(* Schneider Machine Expert - Basic project Projeto Sharpy 2 - Encoder e botão, file version 3.0.0.0 *)
(* ProjectInformations: Name=Novo projeto *)

HARDWARE
  Cpu 0: TM221CE40R
  EthernetConfiguration: NetworkName=M221, IpAllocationMode=FixedAddress, IpAddress=10.0.0.20, SubnetMask=255.0.0.0
  SerialLineConfiguration: Baud=Baud19200, Parity=ParityEven, DataBits=DataBits8, StopBits=StopBits1, PhysicalMedium=PhysicalMediumRs485, TransmissionMode=TransmissionModeModbusRtu, SlaveId=1, Addressing=SlaveAddressing
  MastTask: UsePeriodScanMode=false, PeriodScan=100
  FastTask: Period=255
  CpuBehavior: StartingMode=StartAsPreviousState, AutoSaveRamOnEeprom=true, WatchdogPeriod=250

SYMBOLS  (address, symbol, comment, settings)
  %HSC0.V   VALOR_ENCODER  "Entrada de alta velocidade"
  %S6       SB_TB1S  "Base de tempo de 1 s gerada por um relógio interno"
  %MW0      PULSOS_ENCODER  "Pulsos brutos do encoder"
  %MF2      ANGULO_ATUAL  "Ângulo instantâneo em Graus"
  %MF4      ANGULO_PICO  "Maior ângulo atingido no impacto"
  %MF6      ENERGIA_NOMINAL  "Capacidade da ponta do martelo"
  %MF8      ENERGIA_ABSORVIDA  "Resultado final do ensaio em Joules"
  %MF10     MF_10
  %MF12     MF_12
  %TM0        [Type=TP, Preset=7, Base=OneSecond]
  %TM1        [Type=TP, Preset=7, Base=OneSecond]
  %TM2        [Type=TP, Preset=7, Base=OneSecond]
  %I0.2     BOT_RESET  "Botão físico de zerar encoder e pico"
  %I0.17    SENSOR_PORTA  "Sensor se a porta está fechada"
  %I0.18    SENSOR_BAIXO  "Sensor se o braço está em cima"
  %I0.19    SENSOR_CIMA  "Sensor se o braço está em cima"
  %I0.20    BOTÃO_ZERAR
  %I0.21    BOTÃO_IMPACTO  "Botão que libera para o impacto"
  %I0.22    BOTÃO_DESCER  "Botão que aciona por 7s"
  %I0.23    BOTÃO_SUBIR  "Botão que aciona por 7s"
  %Q0.0       "Motor Descer"
  %Q0.1       "Motor Subir"
  %Q0.2       "Disparo impacto"
  %Q0.3     Q_0_3
  %Q0.4     Q_0_4
  %Q0.5     Q_0_5
  %Q0.14    Q_0_14
  %Q0.15    Q_0_15  "Led porta"
  %IW0.0    IN_ANALOG  "Valor do Potenciômetro"  [Type=Type_0_10V, Scope=Scope_Normal, Minimum=0, Maximum=1000]
  %HSC0       [Type=CounterOrDownCounterBiPhasesX4, Preset=0, DedicatedInputs(DedicatedInput(Activated=true), DedicatedInput(Activated=true)), ReflexOutputs(ReflexOutput(Activated=false, LessThanS0=false, GreaterOrEqualThanS0=false, GreaterOrEqualThanS1=false), ReflexOutput(Activated=false, LessThanS0=false, GreaterOrEqualThanS0=false, GreaterOrEqualThanS1=false)), Thresholds(Threshold(ThresholdType=NotUsed, Pri]

POU Novo POU
  (* SectionNumber=1 *)

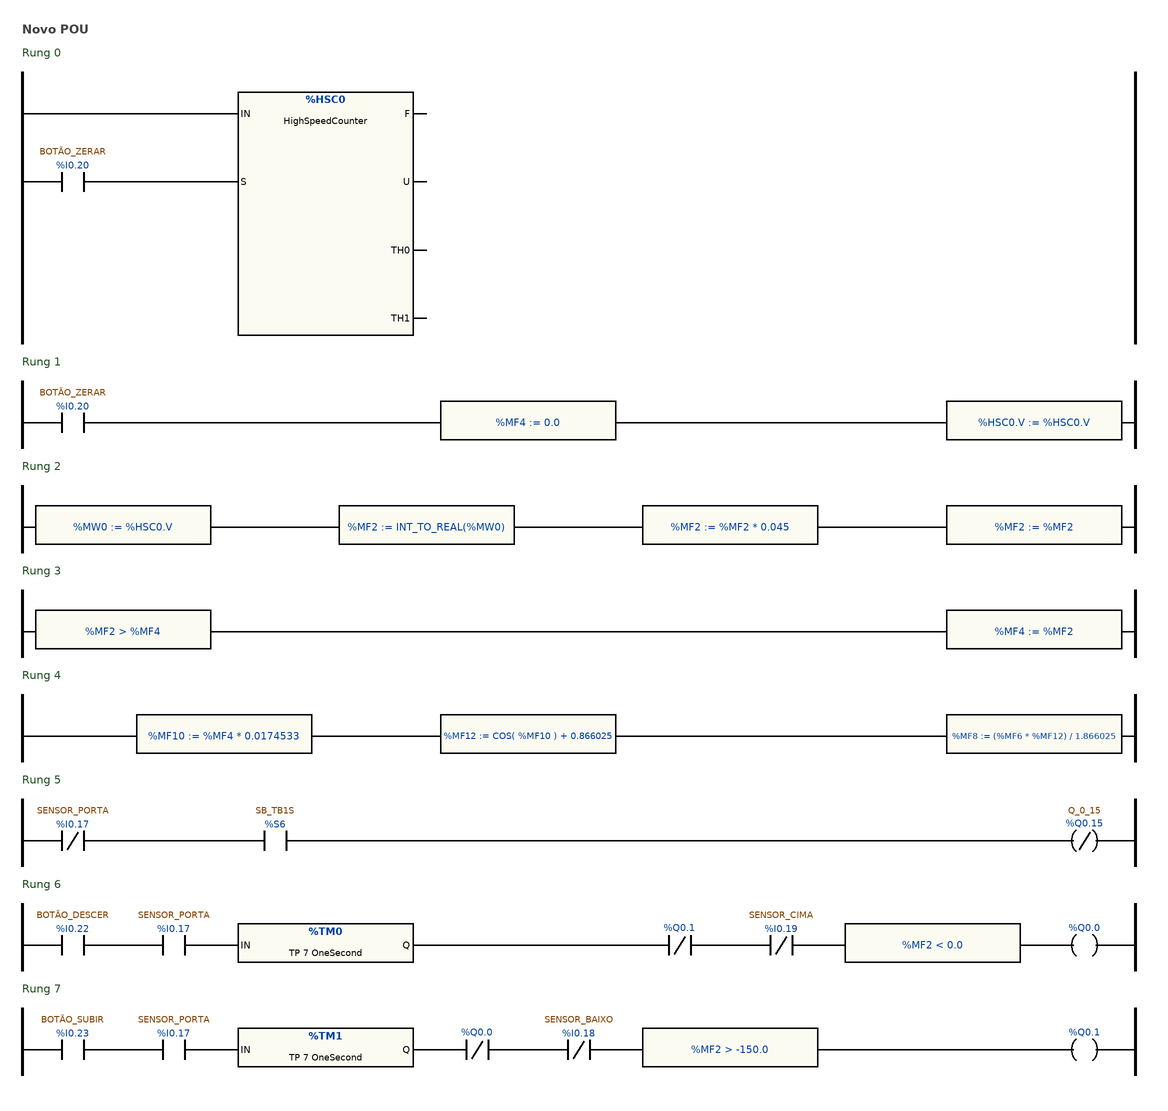

// Rung 0
  BLK %HSC0
  LD 1
  IN
  LD %I0.20               (* BOTÃO_ZERAR *)
  S
  END_BLK
  // as ST:
  //   %HSC0(IN := TRUE, S := BOTÃO_ZERAR);

// Rung 1
  LD %I0.20               (* BOTÃO_ZERAR *)
  OPER [ %MF4 := 0.0 ]    (* ANGULO_PICO *)
  [ %HSC0.V := %HSC0.V ]
  // as ST:
  //   IF BOTÃO_ZERAR THEN ANGULO_PICO := 0.0; END_IF;
  //   IF BOTÃO_ZERAR THEN %HSC0.V := %HSC0.V; END_IF;

// Rung 2
  LD 1
  OPER [ %MW0 := %HSC0.V ](* PULSOS_ENCODER *)
  OPER [ %MF2 := INT_TO_REAL ( %MW0 ) ](* ANGULO_ATUAL, PULSOS_ENCODER *)
  OPER [ %MF2 := %MF2 * 0.045 ](* ANGULO_ATUAL, ANGULO_ATUAL *)
  [ %MF2 := %MF2 ]        (* ANGULO_ATUAL, ANGULO_ATUAL *)
  // as ST:
  //   PULSOS_ENCODER := %HSC0.V;
  //   ANGULO_ATUAL := INT_TO_REAL ( PULSOS_ENCODER );
  //   ANGULO_ATUAL := ANGULO_ATUAL * 0.045;
  //   ANGULO_ATUAL := ANGULO_ATUAL;

// Rung 3
  LD [ %MF2 > %MF4 ]      (* ANGULO_ATUAL, ANGULO_PICO *)
  [ %MF4 := %MF2 ]        (* ANGULO_PICO, ANGULO_ATUAL *)
  // as ST:
  //   IF ANGULO_ATUAL > ANGULO_PICO THEN ANGULO_PICO := ANGULO_ATUAL; END_IF;

// Rung 4
  LD 1
  OPER [ %MF10 := %MF4 * 0.0174533 ](* MF_10, ANGULO_PICO *)
  OPER [ %MF12 := COS ( %MF10 ) + 0.866025 ](* MF_12, MF_10 *)
  [ %MF8 := ( %MF6 * %MF12 ) / 1.866025 ](* ENERGIA_ABSORVIDA, ENERGIA_NOMINAL, MF_12 *)
  // as ST:
  //   MF_10 := ANGULO_PICO * 0.0174533;
  //   MF_12 := COS ( MF_10 ) + 0.866025;
  //   ENERGIA_ABSORVIDA := ( ENERGIA_NOMINAL * MF_12 ) / 1.866025;

// Rung 5
  LDN %I0.17              (* SENSOR_PORTA *)
  AND %S6                 (* SB_TB1S *)
  STN %Q0.15              (* Q_0_15 *)
  // as ST:
  //   Q_0_15 := NOT (NOT SENSOR_PORTA AND SB_TB1S);

// Rung 6
  BLK %TM0
  LD %I0.22               (* BOTÃO_DESCER *)
  AND %I0.17              (* SENSOR_PORTA *)
  IN
  OUT_BLK
  LD Q
  ANDN %Q0.1
  ANDN %I0.19             (* SENSOR_CIMA *)
  AND [ %MF2 < 0.0 ]      (* ANGULO_ATUAL *)
  ST %Q0.0
  END_BLK
  // as ST:
  //   %TM0(IN := BOTÃO_DESCER AND SENSOR_PORTA);
  //   %Q0.0 := %TM0.Q AND NOT %Q0.1 AND NOT SENSOR_CIMA AND ANGULO_ATUAL < 0.0;

// Rung 7
  BLK %TM1
  LD %I0.23               (* BOTÃO_SUBIR *)
  AND %I0.17              (* SENSOR_PORTA *)
  IN
  OUT_BLK
  LD Q
  ANDN %Q0.0
  ANDN %I0.18             (* SENSOR_BAIXO *)
  AND [ %MF2 > -150.0 ]   (* ANGULO_ATUAL *)
  ST %Q0.1
  END_BLK
  // as ST:
  //   %TM1(IN := BOTÃO_SUBIR AND SENSOR_PORTA);
  //   %Q0.1 := %TM1.Q AND NOT %Q0.0 AND NOT SENSOR_BAIXO AND ANGULO_ATUAL > -150.0;

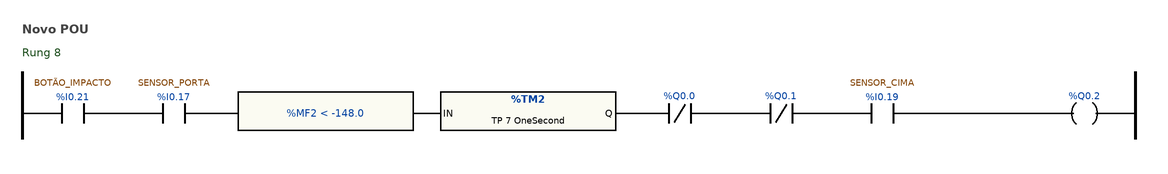

// Rung 8
  BLK %TM2
  LD %I0.21               (* BOTÃO_IMPACTO *)
  AND %I0.17              (* SENSOR_PORTA *)
  AND [ %MF2 < -148.0 ]   (* ANGULO_ATUAL *)
  IN
  OUT_BLK
  LD Q
  ANDN %Q0.0
  ANDN %Q0.1
  AND %I0.19              (* SENSOR_CIMA *)
  ST %Q0.2
  END_BLK
  // as ST:
  //   %TM2(IN := BOTÃO_IMPACTO AND SENSOR_PORTA AND ANGULO_ATUAL < -148.0);
  //   %Q0.2 := %TM2.Q AND NOT %Q0.0 AND NOT %Q0.1 AND SENSOR_CIMA;
